// TIA Portal V20 export
Screen "Pop-up_StyleConfigRFIDRead"  664x479
